(* IEC 61131-3 sources: rusty/tests/lit/single/type_promotion/unary_minus, 5 files *)

(* ---- derived_and_edge_operands.st ---- *)
// RUN: %COMPILE %s && %RUN | %CHECK %s
// A negation of an expression, of a subrange or an enum, and of the smallest LINT, and a negation cut down to a narrow target.
TYPE
    SRU64 : ULINT(0..10);
    SRD : DINT(-10..10);
    EU64 : ULINT (EA := 10, EB := 11);
END_TYPE

VAR_GLOBAL CONSTANT
    csu : SRU64 := 10;
END_VAR

FUNCTION main : DINT
    VAR
        a : USINT := 200;
        s : SINT := -128;
        li : LINT := -9223372036854775808;
        su : SRU64 := 10;
        sd : SRD := -10;
        eu : EU64 := EB;
        d : DINT;
        l : LINT;
        s2 : SINT;
        lr : LREAL;
    END_VAR

    // A negated expression
    d := -(a + 1);
    printf('-(USINT 200 + 1) = %d$N', d);               // CHECK: -(USINT 200 + 1) = -201

    // The smallest LINT has no positive counterpart and wraps to itself
    l := -li;
    printf('-LINT min = %lld$N', l);                    // CHECK-NEXT: -LINT min = -9223372036854775808

    // The DINT result is cut down to a narrow target afterwards
    s2 := -s;
    printf('SINT := -SINT -128 = %d$N', s2);            // CHECK-NEXT: SINT := -SINT -128 = -128

    // A subrange or an enum is negated like its base type, for a variable and for a constant
    lr := -su;
    printf('-SRU64 10 = %.1f$N', lr);                   // CHECK-NEXT: -SRU64 10 = -10.0
    lr := -csu;
    printf('-constant SRU64 10 = %.1f$N', lr);          // CHECK-NEXT: -constant SRU64 10 = -10.0
    d := -sd;
    printf('-SRD -10 = %d$N', d);                       // CHECK-NEXT: -SRD -10 = 10
    l := -eu;
    printf('-EU64 EB = %lld$N', l);                     // CHECK-NEXT: -EU64 EB = -11
END_FUNCTION

(* ---- narrow_operand_widened_to_dint.st ---- *)
// RUN: %COMPILE %s && %RUN | %CHECK %s
// The operand of a negation is widened to DINT first, so a result outside the operand's width does not wrap.
FUNCTION main : DINT
    VAR
        s : SINT := -128;
        i : INT := -32768;
        us : USINT := 200;
        usmax : USINT := 255;
        ui : UINT := 40000;
        uimax : UINT := 65535;
        rd : DINT;
        rl : LINT;
        ri : INT;
    END_VAR

    // Signed minimum values
    rd := -s;
    printf('-SINT -128 = %d$N', rd);        // CHECK: -SINT -128 = 128
    rd := -i;
    printf('-INT -32768 = %d$N', rd);       // CHECK-NEXT: -INT -32768 = 32768

    // Unsigned values above the signed range of the same width
    rd := -us;
    printf('-USINT 200 = %d$N', rd);        // CHECK-NEXT: -USINT 200 = -200
    rd := -usmax;
    printf('-USINT 255 = %d$N', rd);        // CHECK-NEXT: -USINT 255 = -255
    rd := -ui;
    printf('-UINT 40000 = %d$N', rd);       // CHECK-NEXT: -UINT 40000 = -40000
    rd := -uimax;
    printf('-UINT 65535 = %d$N', rd);       // CHECK-NEXT: -UINT 65535 = -65535

    // Typed literal operand
    rd := -USINT#200;
    printf('-USINT#200 = %d$N', rd);        // CHECK-NEXT: -USINT#200 = -200

    // Negation inside a larger expression
    rd := -us + 1;
    printf('-USINT 200 + 1 = %d$N', rd);    // CHECK-NEXT: -USINT 200 + 1 = -199
    printf('-USINT 200 < 0 = %d$N', -us < 0);   // CHECK-NEXT: -USINT 200 < 0 = 1
    printf('-UINT 40000 < 0 = %d$N', -ui < 0);  // CHECK-NEXT: -UINT 40000 < 0 = 1

    // Other targets
    rl := -i;
    printf('LINT := -INT -32768 = %lld$N', rl); // CHECK-NEXT: LINT := -INT -32768 = 32768
    ri := -s;
    printf('INT := -SINT -128 = %d$N', ri);     // CHECK-NEXT: INT := -SINT -128 = 128
END_FUNCTION

(* ---- result_fits_operand_type.st ---- *)
// RUN: %COMPILE %s && %RUN | %CHECK %s
FUNCTION main : DINT
    VAR
        s : SINT := 100;
        i : INT := 30000;
        us : USINT := 100;
        ui : UINT := 30000;
        d : DINT := -2147483647;
        ud : UDINT := 5;
        l : LINT := 9223372036854775807;
        ul : ULINT := 5;
        r : REAL := 1.5;
        rd : DINT;
        rl : LINT;
        rr : REAL;
    END_VAR

    // Narrow operands whose negation fits the operand's width
    rd := -s;
    printf('-SINT 100 = %d$N', rd);         // CHECK: -SINT 100 = -100
    rd := -i;
    printf('-INT 30000 = %d$N', rd);        // CHECK-NEXT: -INT 30000 = -30000
    rd := -us;
    printf('-USINT 100 = %d$N', rd);        // CHECK-NEXT: -USINT 100 = -100
    rd := -ui;
    printf('-UINT 30000 = %d$N', rd);       // CHECK-NEXT: -UINT 30000 = -30000

    // 32-bit and 64-bit operands
    rd := -d;
    printf('-DINT = %d$N', rd);             // CHECK-NEXT: -DINT = 2147483647
    rd := -ud;
    printf('-UDINT 5 = %d$N', rd);          // CHECK-NEXT: -UDINT 5 = -5
    rl := -l;
    printf('-LINT = %lld$N', rl);           // CHECK-NEXT: -LINT = -9223372036854775807
    rl := -ul;
    printf('-ULINT 5 = %lld$N', rl);        // CHECK-NEXT: -ULINT 5 = -5

    // Reals, double negation and the binary form
    rr := -r;
    printf('-REAL 1.5 = %f$N', rr);         // CHECK-NEXT: -REAL 1.5 = -1.500000
    rd := -(-s);
    printf('-(-SINT 100) = %d$N', rd);      // CHECK-NEXT: -(-SINT 100) = 100
    us := 200;
    rd := 0 - us;
    printf('0 - USINT 200 = %d$N', rd);     // CHECK-NEXT: 0 - USINT 200 = -200
END_FUNCTION

(* ---- unsigned_32_bit_operand.st ---- *)
// RUN: %COMPILE %s && %RUN | %CHECK %s
// The negation of a UDINT is LINT, so a value from 2^31 on gives the negative value.
FUNCTION main : DINT
    VAR
        ud : UDINT := 4294967295;
        ud3e9 : UDINT := 3000000000;
        r : LINT;
    END_VAR

    r := -ud;
    printf('-UDINT 4294967295 = %lld$N', r);                // CHECK: -UDINT 4294967295 = -4294967295
    r := -ud3e9;
    printf('-UDINT 3000000000 = %lld$N', r);                // CHECK-NEXT: -UDINT 3000000000 = -3000000000
    printf('-UDINT 3000000000 < 0 = %d$N', -ud3e9 < 0);     // CHECK-NEXT: -UDINT 3000000000 < 0 = 1
END_FUNCTION

(* ---- narrow_constant_widened_to_dint.st ---- *)
// RUN: %COMPILE %s && %RUN | %CHECK %s
// A negated narrow constant is widened to DINT before the negation, so the folded value does not wrap.
VAR_GLOBAL CONSTANT
    cu : USINT := 200;
    ci : INT := -32768;
END_VAR

VAR_GLOBAL
    gu : DINT := -cu;
    gi : DINT := -ci;
END_VAR

PROGRAM prg
    VAR
        mu : DINT := -cu;
    END_VAR
    printf('member := -cu = %d$N', mu);
END_PROGRAM

FUNCTION main : DINT
    VAR CONSTANT
        lc : USINT := 200;
    END_VAR
    VAR
        lu : DINT := -cu;
        rd : DINT;
    END_VAR

    // Global and local initializers
    printf('global := -cu = %d$N', gu);     // CHECK: global := -cu = -200
    printf('global := -ci = %d$N', gi);     // CHECK-NEXT: global := -ci = 32768
    printf('local := -cu = %d$N', lu);      // CHECK-NEXT: local := -cu = -200
    prg();                                  // CHECK-NEXT: member := -cu = -200

    // Body assignments
    rd := -cu;
    printf('body -cu = %d$N', rd);          // CHECK-NEXT: body -cu = -200
    rd := -lc;
    printf('body -lc = %d$N', rd);          // CHECK-NEXT: body -lc = -200
END_FUNCTION
